Staubli VAL3: home.pjx

--- home.pjx ---
Parameters version=s8.15.3Cs9_BS3337 stackSize=5000 millimeterUnit=true
Program file=bind.pgx
Program file=main.pgx
Program file=start.pgx
Program file=stop.pgx
Data file=home.dtx
Library alias=util path=Disk://HMI_cs9/HMI_util/HMI_util.pjx
Library alias=action path=Disk://HMI_cs9/HMI_action/HMI_action.pjx
Library alias=IO path=Disk://HMI_cs9/HMI_IO/HMI_IO.pjx
Library alias=HMI_TRAJ path=Disk://HMI_cs9/HMI_TRAJ/HMI_TRAJ.pjx
Library alias=prog path=Disk://HMI_cs9/HMI_prog/HMI_prog.pjx
Library alias=program path=Disk://source/projectSource/program/program.pjx
Library alias=trajectory path=Disk://source/projectSource/trajectory/trajectory.pjx
Library alias=saveData path=Disk://source/saveData/saveData.pjx
Library alias=HMI_frame path=Disk://HMI_cs9/HMI_FrameSet/HMI_FrameSet.pjx
Library alias=HMI_cycle path=Disk://HMI_cs9/HMI_cycle/HMI_cycle.pjx
Library alias=HMI_setting path=Disk://HMI_cs9/HMI_setting/HMI_setting.pjx
Library alias=HMI_safepoint path=Disk://HMI_cs9/HMI_safepoint/HMI_safepoint.pjx
Library alias=HMI_safezone path=Disk://HMI_cs9/HMI_safezone/HMI_safezone.pjx
Library alias=safecheck path=Disk://source/projectSource/safeCheck/safeCheck.pjx
Library alias=rs path=Disk://source/projectSource/robotStatus/robotStatus.pjx
Library alias=SmartTcp path=Disk://SmartTCP_CS9/SmartTCP_CS9.pjx
Library alias=HMI_message path=Disk://HMI_cs9/HMI_message/HMI_message.pjx

--- home.dtx ---
mdesc mNomSpeed
bool bEditAction
bool bEditIO
bool bEditTRAJ
bool bEditPROG
bool bEditFrame
bool bEditCycle
bool bEditSetting
bool bEditSpoint
bool bEditSzone
string sLib
num nLastStat
string sRobState
bool bExit
public string sVersion
bool bEditTcpTool
bool bLogMsg

--- main.pgx ---
public program main()
  local bool l_bExit
  local bool l_bResult
  local num l_nResult
begin
  util:sPage=""
  do
    if util:sPage!="home"
      util:sPage="home"
      call util:loadingPage()
      call util:initJogMode()


      sLib=toString("",saveData:nLibIndex)
      call bind()
      userPage(util:sPage)
      delay(0.5)
    endIf
    sLib=toString("",saveData:nLibIndex)
    if rs:_nOmacStat!=nLastStat
      nLastStat=rs:_nOmacStat
      if rs:_nOmacStat<9
        userPageAlert("未退出生产模式，主界面按钮锁定！")
        userPageSet("home","btn1","disabled",true)
        userPageSet("home","btn2","disabled",true)
        userPageSet("home","btn3","disabled",true)
        userPageSet("home","btn4","disabled",true)
        userPageSet("home","btn7","disabled",true)
        userPageSet("home","btn8","disabled",true)
        userPageSet("home","btn9","disabled",true)
        userPageSet("home","btn10","disabled",true)
      else
        userPageSet("home","btn1","disabled",false)
        userPageSet("home","btn2","disabled",false)
        userPageSet("home","btn3","disabled",false)
        userPageSet("home","btn4","disabled",false)
        userPageSet("home","btn7","disabled",false)
        userPageSet("home","btn8","disabled",false)
        userPageSet("home","btn9","disabled",false)
        userPageSet("home","btn10","disabled",false)
      endIf
    endIf
    //btn
    if bEditIO
      bEditIO=false
      call IO:main()
    elseIf bEditAction
      bEditAction=false
      call action:main()
    elseIf bEditTRAJ
      bEditTRAJ=false
      call HMI_TRAJ:main()
    elseIf bEditPROG
      bEditPROG=false
      call prog:main()
    elseIf bEditFrame
      bEditFrame=false
      call HMI_frame:main()
    elseIf bEditCycle
      bEditCycle=false
      call HMI_cycle:main()
    elseIf bEditSetting
      bEditSetting=false
      call HMI_setting:main()
    elseIf bEditSpoint
      bEditSpoint=false
      call HMI_safepoint:main()
    elseIf bEditSzone
      bEditSzone=false
      call HMI_safezone:main()
      //guohangxin add 20230323
    elseIf bEditTcpTool
      bEditTcpTool=false
      call util:loadingPage()
      call SmartTcp:start()
      util:sPage=""
    elseIf bLogMsg
      bLogMsg=false
      call HMI_message:main()
    elseIf bExit
      bExit=false
      l_bResult=userPageConfirm("是否退出当前应用？")
      if l_bResult
        rs:bQuitApp=true
      endIf
    endIf

    //rob state
    sRobState=toString(".9",rs:nHWState)
    //jogmode
    call util:jogMode(saveData:nUsingTool,0)
    delay(0)
  until rs:bQuitApp==true
  //rs:bQuitApp=false

end

--- start.pgx ---
program start()
begin
end

--- bind.pgx ---
program bind()
begin
  userPageBindClick("home","btn1",bEditIO,true)
  userPageBindClick("home","btn2",bEditAction,true)
  userPageBindClick("home","btn3",bEditTRAJ,true)
  userPageBindClick("home","btn4",bEditPROG,true)
  userPageBindClick("home","btn7",bEditFrame,true)
  userPageBindClick("home","btn8",bEditSetting,true)
  userPageBindClick("home","btn5",bEditCycle,true)
  userPageBindClick("home","btn6",bLogMsg,true)
  userPageBindClick("home","btn9",bEditSpoint,true)
  userPageBindClick("home","btn10",bEditSzone,true)
  userPageBindClick("home","btn11",bEditTcpTool,true)
  userPageBindClick("home","img1",bExit,true)
  userPageSet("home","btn1","disabled",false)
  userPageSet("home","btn2","disabled",true)
  userPageSet("home","btn3","disabled",false)
  userPageSet("home","btn4","disabled",true)
  userPageSet("home","btn5","disabled",false)
  userPageSet("home","btn6","disabled",false)
  userPageSet("home","btn7","disabled",true)
  userPageSet("home","btn8","disabled",false)
  userPageSet("home","btn9","disabled",true)
  userPageSet("home","btn10","disabled",true)
  userPageSet("home","btn11","disabled",true)

  userPageBind("home","lbl3","innerHTML",sLib,1,"r")
  userPageBind("home","lbl3_Copy1","innerHTML",sRobState,1,"r")
end

--- stop.pgx ---
program stop()
begin
end
